(* IEC 61131-3 sources: SRCI_CLIENT_PLC/RobotLibrary/Library/POUs/General/MC_SwitchLanguage/Structures, 4 files *)

(* ---- SwitchLanguageOutCmd.st ---- *)
{attribute 'pack_mode' := '1'}
// -------------------------------------------------------------------------
//  SRCI Robot Library
// -------------------------------------------------------------------------
//
//  Object:      SwitchLanguageOutCmd
//  Author:      Thorsten Brach
//  Date:        2024-06-30
//
//  Description:
//
//
//  Copyright:
//    (C) 2024 Thorsten Brach. All rights reserved
//             Licensed under the MIT License.
//
//  Disclaimer:
//    This project is provided without any guarantee and can be used for
//    private and commercial purposes. Any use is at the user’s
//    own risk and responsibility.
//
// -------------------------------------------------------------------------
TYPE SwitchLanguageOutCmd :
STRUCT
  /// Two letter code of actual language used at the original operating panel of the robot.
  ActualLanguageCode : STRING(2);
END_STRUCT
END_TYPE

(* ---- SwitchLanguageParCmd.st ---- *)
{attribute 'pack_mode' := '1'}
// -------------------------------------------------------------------------
//  SRCI Robot Library
// -------------------------------------------------------------------------
//
//  Object:      SwitchLanguageParCmd
//  Author:      Thorsten Brach
//  Date:        2024-06-30
//
//  Description:
//
//
//  Copyright:
//    (C) 2024 Thorsten Brach. All rights reserved
//             Licensed under the MIT License.
//
//  Disclaimer:
//    This project is provided without any guarantee and can be used for
//    private and commercial purposes. Any use is at the user’s
//    own risk and responsibility.
//
// -------------------------------------------------------------------------
TYPE SwitchLanguageParCmd :
STRUCT
  /// Two letter code of language to be set at the original operating panel of the robot (default: EN)
  LanguageCode : STRING(2);
END_STRUCT
END_TYPE

(* ---- SwitchLanguageRecvData.st ---- *)
{attribute 'pack_mode' := '1'}
// -------------------------------------------------------------------------
//  SRCI Robot Library
// -------------------------------------------------------------------------
//
//  Object:      SwitchLanguageRecvData
//  Author:      Thorsten Brach
//  Date:        2024-06-30
//
//  Description:
//
//
//  Copyright:
//    (C) 2024 Thorsten Brach. All rights reserved
//             Licensed under the MIT License.
//
//  Disclaimer:
//    This project is provided without any guarantee and can be used for
//    private and commercial purposes. Any use is at the user’s
//    own risk and responsibility.
//
// -------------------------------------------------------------------------
TYPE SwitchLanguageRecvData EXTENDS RspHeader :
STRUCT
  /// Two letter code of actual language used at the original operating panel of the robot.
  ActualLanguageCode : STRING(2);
END_STRUCT
END_TYPE

(* ---- SwitchLanguageSendData.st ---- *)
{attribute 'pack_mode' := '1'}
// -------------------------------------------------------------------------
//  SRCI Robot Library
// -------------------------------------------------------------------------
//
//  Object:      SwitchLanguageSendData
//  Author:      Thorsten Brach
//  Date:        2024-06-30
//
//  Description:
//
//
//  Copyright:
//    (C) 2024 Thorsten Brach. All rights reserved
//             Licensed under the MIT License.
//
//  Disclaimer:
//    This project is provided without any guarantee and can be used for
//    private and commercial purposes. Any use is at the user’s
//    own risk and responsibility.
//
// -------------------------------------------------------------------------
TYPE SwitchLanguageSendData EXTENDS CmdHeader:
STRUCT
  /// Two letter code of language to be set at the original operating panel of the robot (default: EN)
  LanguageCode : STRING(2);
END_STRUCT
END_TYPE
